{attribute 'qualified_only'}
{attribute 'strict'}
TYPE E_SkidZone :
(
	eCIP := 0,
	eTriBlender,
	eMarinade,
	eColor,
	eLast
);
END_TYPE

(* stored: Version 1.1.0.1, ProductVersion 3.1.4024.15
   DUT E_SkidZone: Id {aa405c71-53c2-4cc6-9ffc-e3f9e6d768b0} *)
